// TwinCAT 3 PLC project EventFramework
// Title: EventFramework
// Company: DM
// ProjectVersion: 1.0.0.2
// Description: Text-list driven alarms and messages on top of Tc3_EventLogger.
// ProgramVersion: 3.1.4026.26
// libraries:
//   Tc2_Standard, * (Beckhoff Automation GmbH)
//   Tc2_System, * (Beckhoff Automation GmbH)
//   Tc3_EventLogger, * (Beckhoff Automation GmbH)
// project tree:
//   DUTs/ E_Language.TcDUT, ST_EventDefinition.TcDUT
//   / GVL_EventDefaults.TcGVL, GVL_EventFramework.TcGVL
//   Interfaces/ I_Alarm.TcIO, I_ArgumentBuilder.TcIO, I_ArgumentSource.TcIO, I_CatalogEvent.TcIO, I_EventContext.TcIO, I_EventEntryProvider.TcIO, I_LanguageProvider.TcIO, I_Message.TcIO, I_TextFormatter.TcIO, I_TextProvider.TcIO
//   POUs/ FB_CatalogAlarm.TcPOU, FB_CatalogEventBase.TcPOU, FB_CatalogMessage.TcPOU, FB_DefinitionTextProvider.TcPOU, FB_EventArgs.TcPOU, FB_EventContext.TcPOU, FB_GenericEventClass.TcPOU, FB_LanguageSelector.TcPOU, FB_PlaceholderFormatter.TcPOU
// (motion and I/O tree: see PLC project eventloggersample)
// real-time tasks:
//   TASK PlcTask: cycle T#10ms, priority 20, ADS port 350

// ---- DUTs/E_Language.TcDUT
// Languages of the event texts. The first value is the default/fallback language.
// Adding one: add a value here, raise GVL_EventFramework.cLanguageCount,
// then add the translation to the lines in GVL_EventTexts (missing ones fall back to the default).
// Only languages whose characters fit in STRING (Windows-1252); other alphabets would need WSTRING.
{attribute 'qualified_only'}
TYPE E_Language :
(
	English		:= 0,
	German		:= 1,
	French		:= 2,
	Spanish		:= 3,
	Italian		:= 4,
	Portuguese	:= 5,
	Dutch		:= 6,
	Danish		:= 7,
	Swedish		:= 8,
	Norwegian	:= 9,
	Finnish		:= 10
) USINT;
END_TYPE

// ---- DUTs/ST_EventDefinition.TcDUT
// One event of the text list (see GVL_EventTexts).
TYPE ST_EventDefinition :
STRUCT
	nId					: UDINT;			// stable key: source info nId, HMI filtering, external (CSV) texts
	eSeverity			: TcEventSeverity;	// selects the generic TMC event (Verbose/Info/Warning/Error/Critical)
	bWithConfirmation	: BOOL;				// alarms only: operator has to confirm
	asText				: ARRAY[0..GVL_EventFramework.cLanguageCount - 1] OF STRING(160);	// per E_Language, {0}..{9} = arguments
END_STRUCT
END_TYPE

// ---- GVL_EventDefaults.TcGVL
// Default composition root: used by every catalog event that has no Context of its own.
// Fully wired: an application needs no setup of its own.
// Replace any part at startup, e.g.  GVL_EventDefaults.fbContext.Texts := fbCsvTexts;
{attribute 'qualified_only'}
VAR_GLOBAL
	fbDefinitionTexts	: FB_DefinitionTextProvider;
	fbLanguage			: FB_LanguageSelector;
	fbFormatter			: FB_PlaceholderFormatter;
	fbEventClass		: FB_GenericEventClass;
	fbContext			: FB_EventContext(ipTexts := fbDefinitionTexts,
										  ipLanguage := fbLanguage,
										  ipFormatter := fbFormatter,
										  ipEventEntries := fbEventClass);
END_VAR

// ---- GVL_EventFramework.TcGVL
{attribute 'qualified_only'}
VAR_GLOBAL CONSTANT
	cMaxArguments		: USINT := 10;				// placeholders {0}..{9}
	cLanguageCount		: USINT := 11;				// number of values in E_Language - raise when adding a language
	HR_NO_CONTEXT		: HRESULT := -2147467261;	// 16#80004003 (E_POINTER): no I_EventContext was injected
	HR_NOT_IMPLEMENTED	: HRESULT := -2147467263;	// 16#80004001 (E_NOTIMPL)
END_VAR

// ---- Interfaces/I_Alarm.TcIO
INTERFACE I_Alarm EXTENDS I_CatalogEvent

METHOD Raise : HRESULT
END_METHOD

METHOD Clear : HRESULT
VAR_INPUT
	bResetConfirmation	: BOOL;
END_VAR
END_METHOD

METHOD Confirm : HRESULT
END_METHOD

// Level driven: raises while bActive is TRUE, clears when it drops.
METHOD SetActive : HRESULT
VAR_INPUT
	bActive	: BOOL;
END_VAR
END_METHOD

PROPERTY IsRaised : BOOL
GET
END_GET
END_PROPERTY

PROPERTY ConfirmationState : TcEventConfirmationState
GET
END_GET
END_PROPERTY

END_INTERFACE

// ---- Interfaces/I_ArgumentBuilder.TcIO
// Write side of the event arguments (fluent).
INTERFACE I_ArgumentBuilder

METHOD Clear : I_ArgumentBuilder
END_METHOD

METHOD AddString : I_ArgumentBuilder
VAR_INPUT
	sValue	: T_MaxString;
END_VAR
END_METHOD

METHOD AddDInt : I_ArgumentBuilder
VAR_INPUT
	nValue	: DINT;
END_VAR
END_METHOD

METHOD AddLReal : I_ArgumentBuilder
VAR_INPUT
	fValue		: LREAL;
	nDecimals	: USINT;	// 0..9
END_VAR
END_METHOD

METHOD AddBool : I_ArgumentBuilder
VAR_INPUT
	bValue	: BOOL;
END_VAR
END_METHOD

END_INTERFACE

// ---- Interfaces/I_ArgumentSource.TcIO
// Read side of the event arguments (used by formatters).
INTERFACE I_ArgumentSource

PROPERTY Count : USINT
GET
END_GET
END_PROPERTY

METHOD GetArgument : T_MaxString
VAR_INPUT
	nIndex	: USINT;
END_VAR
END_METHOD

END_INTERFACE

// ---- Interfaces/I_CatalogEvent.TcIO
// Common part of catalog alarms and messages.
INTERFACE I_CatalogEvent

PROPERTY Arguments : I_ArgumentBuilder
GET
END_GET
END_PROPERTY

PROPERTY Severity : TcEventSeverity
GET
END_GET
END_PROPERTY

PROPERTY LastResult : HRESULT
GET
END_GET
END_PROPERTY

PROPERTY SourceName : T_MaxString
GET
END_GET
SET
END_SET
END_PROPERTY

END_INTERFACE

// ---- Interfaces/I_EventContext.TcIO
// Bundles the services every catalog event needs (injected once).
INTERFACE I_EventContext

PROPERTY Texts : I_TextProvider
GET
END_GET
END_PROPERTY

PROPERTY Language : I_LanguageProvider
GET
END_GET
END_PROPERTY

PROPERTY Formatter : I_TextFormatter
GET
END_GET
END_PROPERTY

PROPERTY EventEntries : I_EventEntryProvider
GET
END_GET
END_PROPERTY

END_INTERFACE

// ---- Interfaces/I_EventEntryProvider.TcIO
// Maps a severity onto a TMC event (event class + event id).
INTERFACE I_EventEntryProvider

METHOD GetEventEntry : TcEventEntry
VAR_INPUT
	eSeverity	: TcEventSeverity;
END_VAR
END_METHOD

END_INTERFACE

// ---- Interfaces/I_LanguageProvider.TcIO
// Current language of the event texts.
INTERFACE I_LanguageProvider

PROPERTY Current : E_Language
GET
END_GET
END_PROPERTY

END_INTERFACE

// ---- Interfaces/I_Message.TcIO
INTERFACE I_Message EXTENDS I_CatalogEvent

METHOD Send : HRESULT
END_METHOD

END_INTERFACE

// ---- Interfaces/I_TextFormatter.TcIO
// Renders a text template with arguments.
INTERFACE I_TextFormatter

METHOD Format : T_MaxString
VAR_INPUT
	ipArguments	: I_ArgumentSource;
END_VAR
VAR_IN_OUT CONSTANT
	sTemplate	: T_MaxString;
END_VAR
END_METHOD

END_INTERFACE

// ---- Interfaces/I_TextProvider.TcIO
// Supplies the text template of an event in a language.
// Default: FB_DefinitionTextProvider (texts from GVL_EventTexts).
// Extension point: e.g. a CSV provider that overrides texts and delegates to the default.
INTERFACE I_TextProvider

METHOD GetTemplate : T_MaxString
VAR_INPUT
	eLanguage		: E_Language;
END_VAR
VAR_IN_OUT CONSTANT
	stDefinition	: ST_EventDefinition;
END_VAR
END_METHOD

END_INTERFACE

// ---- POUs/FB_DefinitionTextProvider.TcPOU
// Default I_TextProvider: takes the text from the definition itself (GVL_EventTexts).
// Falls back to the default language (index 0) when a translation is missing.
FUNCTION_BLOCK FB_DefinitionTextProvider IMPLEMENTS I_TextProvider
VAR
END_VAR

METHOD GetTemplate : T_MaxString
VAR_INPUT
	eLanguage		: E_Language;
END_VAR
VAR_IN_OUT CONSTANT
	stDefinition	: ST_EventDefinition;
END_VAR
VAR
	nIndex	: USINT;
END_VAR
nIndex := eLanguage;
IF nIndex < GVL_EventFramework.cLanguageCount AND_THEN LEN(stDefinition.asText[nIndex]) > 0 THEN
	GetTemplate := stDefinition.asText[nIndex];
ELSE
	GetTemplate := stDefinition.asText[0];
END_IF
END_METHOD

END_FUNCTION_BLOCK

// ---- POUs/FB_LanguageSelector.TcPOU
// Holds the current event text language. Affects events raised after the change.
FUNCTION_BLOCK FB_LanguageSelector IMPLEMENTS I_LanguageProvider
VAR
	_eCurrent	: E_Language;
END_VAR

PROPERTY Current : E_Language
GET
Current := _eCurrent;
END_GET
SET
_eCurrent := Current;
END_SET
END_PROPERTY

END_FUNCTION_BLOCK

// ---- POUs/FB_PlaceholderFormatter.TcPOU
// Replaces {0}..{9} in a template with the matching argument.
// Placeholders without an argument are left in the text so they are easy to spot.
FUNCTION_BLOCK FB_PlaceholderFormatter IMPLEMENTS I_TextFormatter
VAR
END_VAR

METHOD Format : T_MaxString
VAR_INPUT
	ipArguments	: I_ArgumentSource;
END_VAR
VAR_IN_OUT CONSTANT
	sTemplate	: T_MaxString;
END_VAR
VAR
	sResult			: T_MaxString;
	sArgument		: T_MaxString;
	nLen			: INT;
	nIn				: INT;
	nOut			: INT;
	nArg			: INT;
	nArgLen			: INT;
	nIndex			: USINT;
	bPlaceholder	: BOOL;
END_VAR
VAR CONSTANT
	cOpen		: BYTE := 16#7B;	// {
	cClose		: BYTE := 16#7D;	// }
	cZero		: BYTE := 16#30;	// 0
	cNine		: BYTE := 16#39;	// 9
	cMaxLen		: INT := 255;
END_VAR
nLen := LEN(sTemplate);

WHILE nIn < nLen AND nOut < cMaxLen DO
	bPlaceholder := FALSE;
	IF nIn + 2 < nLen
		AND_THEN sTemplate[nIn] = cOpen
		AND_THEN sTemplate[nIn + 1] >= cZero
		AND_THEN sTemplate[nIn + 1] <= cNine
		AND_THEN sTemplate[nIn + 2] = cClose
		AND_THEN ipArguments <> 0
	THEN
		nIndex := BYTE_TO_USINT(sTemplate[nIn + 1] - cZero);
		bPlaceholder := nIndex < ipArguments.Count;
	END_IF

	IF bPlaceholder THEN
		sArgument := ipArguments.GetArgument(nIndex);
		nArgLen := LEN(sArgument);
		nArg := 0;
		WHILE nArg < nArgLen AND nOut < cMaxLen DO
			sResult[nOut] := sArgument[nArg];
			nOut := nOut + 1;
			nArg := nArg + 1;
		END_WHILE
		nIn := nIn + 3;
	ELSE
		sResult[nOut] := sTemplate[nIn];
		nOut := nOut + 1;
		nIn := nIn + 1;
	END_IF
END_WHILE

sResult[nOut] := 0;
Format := sResult;
END_METHOD

END_FUNCTION_BLOCK

// ---- POUs/FB_GenericEventClass.TcPOU
// The ONLY place that knows the TMC event class "GenericEvents".
// Each event in that class has the text "{0}", the full text is supplied as argument.
// The class is pinned in this library (Add > Global Data Type), so it is added to the
// type system of every project that references the library.
// Used by GVL_EventDefaults.fbContext.
FUNCTION_BLOCK FB_GenericEventClass IMPLEMENTS I_EventEntryProvider
VAR
END_VAR

METHOD GetEventEntry : TcEventEntry
VAR_INPUT
	eSeverity	: TcEventSeverity;
END_VAR
CASE eSeverity OF
	TcEventSeverity.Verbose:	GetEventEntry := TC_EVENTS.GenericEvents.Verbose;
	TcEventSeverity.Info:		GetEventEntry := TC_EVENTS.GenericEvents.Info;
	TcEventSeverity.Warning:	GetEventEntry := TC_EVENTS.GenericEvents.Warning;
	TcEventSeverity.Error:		GetEventEntry := TC_EVENTS.GenericEvents.Error;
	TcEventSeverity.Critical:	GetEventEntry := TC_EVENTS.GenericEvents.Critical;
ELSE
	GetEventEntry := TC_EVENTS.GenericEvents.Error;
END_CASE
END_METHOD

END_FUNCTION_BLOCK

// ---- POUs/FB_EventContext.TcPOU
// Composition of the event services, built once in a composition root (see GVL_EventDefaults).
// The setters let an application swap a single service; set them before the first event is raised.
FUNCTION_BLOCK FB_EventContext IMPLEMENTS I_EventContext
VAR
	_ipTexts		: I_TextProvider;
	_ipLanguage		: I_LanguageProvider;
	_ipFormatter	: I_TextFormatter;
	_ipEventEntries	: I_EventEntryProvider;
END_VAR

METHOD FB_init : BOOL
VAR_INPUT
	bInitRetains	: BOOL;
	bInCopyCode		: BOOL;
	ipTexts			: I_TextProvider;
	ipLanguage		: I_LanguageProvider;
	ipFormatter		: I_TextFormatter;
	ipEventEntries	: I_EventEntryProvider;
END_VAR
_ipTexts := ipTexts;
_ipLanguage := ipLanguage;
_ipFormatter := ipFormatter;
_ipEventEntries := ipEventEntries;
END_METHOD

PROPERTY Texts : I_TextProvider
GET
Texts := _ipTexts;
END_GET
SET
_ipTexts := Texts;
END_SET
END_PROPERTY

PROPERTY Language : I_LanguageProvider
GET
Language := _ipLanguage;
END_GET
SET
_ipLanguage := Language;
END_SET
END_PROPERTY

PROPERTY Formatter : I_TextFormatter
GET
Formatter := _ipFormatter;
END_GET
SET
_ipFormatter := Formatter;
END_SET
END_PROPERTY

PROPERTY EventEntries : I_EventEntryProvider
GET
EventEntries := _ipEventEntries;
END_GET
SET
_ipEventEntries := EventEntries;
END_SET
END_PROPERTY

END_FUNCTION_BLOCK

// ---- POUs/FB_CatalogAlarm.TcPOU
// Stateful alarm whose severity and text come from the event catalog.
// Declare as:  fbX : FB_CatalogAlarm(stDefinition := GVL_EventTexts.X);
FUNCTION_BLOCK FB_CatalogAlarm EXTENDS FB_CatalogEventBase IMPLEMENTS I_Alarm
VAR
	_fbAlarm	: FB_TcAlarm;
END_VAR

METHOD PROTECTED CreateEvent : HRESULT
VAR_INPUT
	stEventEntry	: TcEventEntry;
	ipSourceInfo	: I_TcSourceInfo;
END_VAR
CreateEvent := _fbAlarm.CreateEx(stEventEntry := stEventEntry,
								 bWithConfirmation := _stDefinition.bWithConfirmation,
								 ipSourceInfo := ipSourceInfo);
END_METHOD

METHOD Raise : HRESULT
VAR
	sText	: T_MaxString;
END_VAR
IF NOT EnsureCreated() THEN
	Raise := _hrLast;
	RETURN;
END_IF

// Already active: keep the original text and timestamp
IF _fbAlarm.bRaised THEN
	RETURN;
END_IF

sText := BuildText();
_fbAlarm.ipArguments.Clear().AddString(sText);
_hrLast := _fbAlarm.Raise(0);
Raise := _hrLast;
END_METHOD

METHOD Clear : HRESULT
VAR_INPUT
	bResetConfirmation	: BOOL;
END_VAR
IF NOT _bCreated THEN
	RETURN;
END_IF
_hrLast := _fbAlarm.Clear(0, bResetConfirmation);
Clear := _hrLast;
END_METHOD

METHOD Confirm : HRESULT
IF NOT _bCreated THEN
	RETURN;
END_IF
_hrLast := _fbAlarm.Confirm(0);
Confirm := _hrLast;
END_METHOD

METHOD SetActive : HRESULT
VAR_INPUT
	bActive	: BOOL;
END_VAR
IF bActive AND NOT IsRaised THEN
	SetActive := Raise();
ELSIF NOT bActive AND IsRaised THEN
	SetActive := Clear(bResetConfirmation := FALSE);
END_IF
END_METHOD

PROPERTY IsRaised : BOOL
GET
IsRaised := _bCreated AND_THEN _fbAlarm.bRaised;
END_GET
END_PROPERTY

PROPERTY ConfirmationState : TcEventConfirmationState
GET
ConfirmationState := _fbAlarm.eConfirmationState;
END_GET
END_PROPERTY

END_FUNCTION_BLOCK

// ---- POUs/FB_CatalogEventBase.TcPOU
// Shared behaviour of catalog alarms and messages:
//  - gets its definition (severity, confirmation, texts) from GVL_EventTexts at declaration
//  - owns a unique source info (default name = instance path, nId = definition nId),
//    so any number of catalog events can be active at the same time even when
//    they map onto the same generic TMC event
//  - gets the text in the current language and renders it with the context's formatter
//  - uses GVL_EventDefaults.fbContext unless another context is set via Context
// Derived blocks only create/drive their concrete Tc3_EventLogger object.
{attribute 'reflection'}
FUNCTION_BLOCK ABSTRACT FB_CatalogEventBase IMPLEMENTS I_CatalogEvent
VAR
	{attribute 'instance-path'}
	{attribute 'noinit'}
	_sInstancePath	: T_MaxString;
END_VAR
VAR
	_ipContext		: I_EventContext;		// 0 = GVL_EventDefaults.fbContext
	_stDefinition	: ST_EventDefinition;
	_fbSourceInfo	: FB_TcSourceInfo;
	_fbArguments	: FB_EventArgs;
	_sSourceName	: T_MaxString;
	_bCreated		: BOOL;
	_hrLast			: HRESULT;
END_VAR

METHOD FB_init : BOOL
VAR_INPUT
	bInitRetains	: BOOL;
	bInCopyCode		: BOOL;
	stDefinition	: ST_EventDefinition;	// e.g. GVL_EventTexts.ConveyorJam
END_VAR
_stDefinition := stDefinition;
END_METHOD

// Lazily creates the event logger object on first use.
METHOD PROTECTED EnsureCreated : BOOL
VAR
	ipContext	: I_EventContext;
	ipEntries	: I_EventEntryProvider;
END_VAR
IF _bCreated THEN
	EnsureCreated := TRUE;
	RETURN;
END_IF

ipContext := Context;
IF ipContext = 0 THEN
	_hrLast := GVL_EventFramework.HR_NO_CONTEXT;
	RETURN;
END_IF

// No TMC mapping (only possible when a custom context leaves EventEntries empty)
ipEntries := ipContext.EventEntries;
IF ipEntries = 0 THEN
	_hrLast := GVL_EventFramework.HR_NO_CONTEXT;
	RETURN;
END_IF

// Unique source info per instance => simultaneous events never collide
IF _sSourceName = '' THEN
	_sSourceName := _sInstancePath;
END_IF
_fbSourceInfo.sName := _sSourceName;
_fbSourceInfo.nId := _stDefinition.nId;

_hrLast := CreateEvent(stEventEntry := ipEntries.GetEventEntry(_stDefinition.eSeverity),
					   ipSourceInfo := _fbSourceInfo);
_bCreated := SUCCEEDED(_hrLast);
EnsureCreated := _bCreated;
END_METHOD

// Template method: derived blocks create their FB_TcAlarm / FB_TcMessage here.
METHOD PROTECTED CreateEvent : HRESULT
VAR_INPUT
	stEventEntry	: TcEventEntry;
	ipSourceInfo	: I_TcSourceInfo;
END_VAR
CreateEvent := GVL_EventFramework.HR_NOT_IMPLEMENTED;
END_METHOD

// Template in the current language, placeholders replaced by the arguments.
METHOD PROTECTED BuildText : T_MaxString
VAR
	ipContext	: I_EventContext;
	ipTexts		: I_TextProvider;
	ipLanguage	: I_LanguageProvider;
	ipFormatter	: I_TextFormatter;
	eLanguage	: E_Language;
	sTemplate	: T_MaxString;
END_VAR
ipContext := Context;
ipTexts := ipContext.Texts;
ipLanguage := ipContext.Language;
ipFormatter := ipContext.Formatter;

IF ipLanguage <> 0 THEN
	eLanguage := ipLanguage.Current;
END_IF

IF ipTexts <> 0 THEN
	sTemplate := ipTexts.GetTemplate(eLanguage := eLanguage, stDefinition := _stDefinition);
ELSE
	sTemplate := _stDefinition.asText[0];
END_IF
IF sTemplate = '' THEN
	sTemplate := CONCAT('Event ', UDINT_TO_STRING(_stDefinition.nId));
END_IF

IF ipFormatter <> 0 THEN
	BuildText := ipFormatter.Format(ipArguments := _fbArguments, sTemplate := sTemplate);
ELSE
	BuildText := sTemplate;
END_IF
END_METHOD

// Arguments are taken over when the event is raised/sent.
PROPERTY Arguments : I_ArgumentBuilder
GET
Arguments := _fbArguments;
END_GET
END_PROPERTY

// Event services used by this event (default: GVL_EventDefaults.fbContext).
// Set it only to inject a different context; only effective before the first Raise/Send.
PROPERTY Context : I_EventContext
GET
IF _ipContext <> 0 THEN
	Context := _ipContext;
ELSE
	Context := GVL_EventDefaults.fbContext;
END_IF
END_GET
SET
IF NOT _bCreated THEN
	_ipContext := Context;
END_IF
END_SET
END_PROPERTY

PROPERTY Severity : TcEventSeverity
GET
Severity := _stDefinition.eSeverity;
END_GET
END_PROPERTY

PROPERTY LastResult : HRESULT
GET
LastResult := _hrLast;
END_GET
END_PROPERTY

// Optional override of the source name (default: instance path).
// Only effective before the first Raise/Send.
PROPERTY SourceName : T_MaxString
GET
SourceName := _sSourceName;
END_GET
SET
IF NOT _bCreated THEN
	_sSourceName := SourceName;
END_IF
END_SET
END_PROPERTY

END_FUNCTION_BLOCK

// ---- POUs/FB_EventArgs.TcPOU
// Argument container. Values are stored as text, ready for the formatter.
FUNCTION_BLOCK FB_EventArgs IMPLEMENTS I_ArgumentBuilder, I_ArgumentSource
VAR
	aValues	: ARRAY[0..GVL_EventFramework.cMaxArguments - 1] OF T_MaxString;
	nCount	: USINT;
END_VAR

METHOD PRIVATE Append : I_ArgumentBuilder
VAR_INPUT
	sValue	: T_MaxString;
END_VAR
IF nCount < GVL_EventFramework.cMaxArguments THEN
	aValues[nCount] := sValue;
	nCount := nCount + 1;
END_IF
Append := THIS^;
END_METHOD

METHOD Clear : I_ArgumentBuilder
nCount := 0;
Clear := THIS^;
END_METHOD

METHOD AddString : I_ArgumentBuilder
VAR_INPUT
	sValue	: T_MaxString;
END_VAR
AddString := Append(sValue);
END_METHOD

METHOD AddDInt : I_ArgumentBuilder
VAR_INPUT
	nValue	: DINT;
END_VAR
AddDInt := Append(DINT_TO_STRING(nValue));
END_METHOD

METHOD AddLReal : I_ArgumentBuilder
VAR_INPUT
	fValue		: LREAL;
	nDecimals	: USINT;	// 0..9
END_VAR
VAR
	nDigits	: USINT;
	nScale	: LINT := 1;
	nScaled	: LINT;
	i		: USINT;
	sFrac	: STRING(20);
	sValue	: T_MaxString;
END_VAR
nDigits := MIN(nDecimals, 9);
FOR i := 1 TO nDigits DO
	nScale := nScale * 10;
END_FOR

// Fixed-point formatting avoids LREAL_TO_STRING artefacts like 82.350000000000009
nScaled := LREAL_TO_LINT(ABS(fValue) * LINT_TO_LREAL(nScale));
sValue := LINT_TO_STRING(nScaled / nScale);
IF nDigits > 0 THEN
	sFrac := LINT_TO_STRING(nScaled MOD nScale);
	WHILE LEN(sFrac) < nDigits DO
		sFrac := CONCAT('0', sFrac);
	END_WHILE
	sValue := CONCAT(CONCAT(sValue, '.'), sFrac);
END_IF
IF fValue < 0 AND nScaled <> 0 THEN
	sValue := CONCAT('-', sValue);
END_IF

AddLReal := Append(sValue);
END_METHOD

METHOD AddBool : I_ArgumentBuilder
VAR_INPUT
	bValue	: BOOL;
END_VAR
IF bValue THEN
	AddBool := Append('TRUE');
ELSE
	AddBool := Append('FALSE');
END_IF
END_METHOD

METHOD GetArgument : T_MaxString
VAR_INPUT
	nIndex	: USINT;
END_VAR
IF nIndex < nCount THEN
	GetArgument := aValues[nIndex];
END_IF
END_METHOD

PROPERTY Count : USINT
GET
Count := nCount;
END_GET
END_PROPERTY

END_FUNCTION_BLOCK

// ---- POUs/FB_CatalogMessage.TcPOU
// Fire-and-forget message whose severity and text come from the event catalog.
FUNCTION_BLOCK FB_CatalogMessage EXTENDS FB_CatalogEventBase IMPLEMENTS I_Message
VAR
	_fbMessage	: FB_TcMessage;
END_VAR

METHOD PROTECTED CreateEvent : HRESULT
VAR_INPUT
	stEventEntry	: TcEventEntry;
	ipSourceInfo	: I_TcSourceInfo;
END_VAR
CreateEvent := _fbMessage.CreateEx(stEventEntry := stEventEntry, ipSourceInfo := ipSourceInfo);
END_METHOD

METHOD Send : HRESULT
VAR
	sText	: T_MaxString;
END_VAR
IF NOT EnsureCreated() THEN
	Send := _hrLast;
	RETURN;
END_IF

sText := BuildText();
_fbMessage.ipArguments.Clear().AddString(sText);
_hrLast := _fbMessage.Send(0);
Send := _hrLast;
END_METHOD

END_FUNCTION_BLOCK
